(* IEC 61131-3 sources: ControlsBenchMUSE/codesys/demo/source, 10 files *)

(* ---- ST_BenchInputImage.st ---- *)
TYPE ST_BenchInputImage :
STRUCT
    PE_Entry : BOOL;
    PE_D1Approach : BOOL;
    PE_D2Approach : BOOL;
    PE_ExitA : BOOL;
    PE_ExitB : BOOL;
    PE_Runout : BOOL;
    D1_HomeFB : BOOL;
    D1_ExtendedFB : BOOL;
    D2_HomeFB : BOOL;
    D2_ExtendedFB : BOOL;
    Drive_RunningFB : BOOL;
    Drive_Overload : BOOL;
    ExitA_Ready : BOOL;
    ExitB_Ready : BOOL;
    Runout_Ready : BOOL;
    Belt_SpeedActual : REAL;
    Drive_Current : REAL;
    D1_Position : REAL;
    D2_Position : REAL;
    Encoder_Count : UDINT;
END_STRUCT
END_TYPE

(* ---- ST_DemoStatus.st ---- *)
TYPE ST_DemoStatus :
STRUCT
    Mode : UINT;
    ModeText : STRING(16);
    FaultCode : UINT;
    FaultText : STRING(80);
    ExceptionCode : UINT;
    ExceptionText : STRING(80);
    Motor_RunCmd : BOOL;
    D1_ExtendCmd : BOOL;
    D2_ExtendCmd : BOOL;
    StackLight_Red : BOOL;
    StackLight_Green : BOOL;
    ReleaseReady : BOOL;
    ItemActive : BOOL;
    ActiveItemId : UDINT;
    RequestedRoute : UINT;
    EffectiveRoute : UINT;
    ActualExit : UINT;
    Disposition : UINT;
    OfferAckSequence : UDINT;
    OfferAckItemId : UDINT;
    OfferAccepted : BOOL;
    OfferReason : UINT;
    OfferPending : BOOL;
    CompletionSequence : UDINT;
    CompletionPending : BOOL;
    CompletionItemId : UDINT;
    CompletionRoute : UINT;
    CompletionExit : UINT;
    CompletionDisposition : UINT;
    CountExitA : UDINT;
    CountExitB : UDINT;
    CountRunout : UDINT;
    CountMisroute : UDINT;
    CountFaulted : UDINT;
    StartAck : UDINT;
    StopAck : UDINT;
    ResetAck : UDINT;
    StartAccepted : BOOL;
    ResetAccepted : BOOL;
    EncoderDelta : UDINT;
    BeltSpeedMps : LREAL;
    TravelMetres : LREAL;
    ScanTimeUs : ULINT;
END_STRUCT
END_TYPE

(* ---- GVL_BenchRead.st ---- *)
NAMESPACE GVL_BenchRead
{attribute 'qualified_only'}
VAR_GLOBAL
    // Bench state and liveness. Workstation read-only through OPC UA.
    SimApplied : BOOL := FALSE;
    ConnectorStale : BOOL := TRUE;
    ActiveSlot : USINT := 255;
    AppliedEpoch : ULINT := 0;
    AppliedSequence : ULINT := 0;
    // Published compatibility placeholders retained by the configured symbol type.
    AppliedCaptureCycle : ULINT := 0;
    AppliedCaptureTimeUs : ULINT := 0;
    PlcHeartbeat : ULINT := 0;
    PlcBootIdentity : ULINT := 0;
    PlcCycle : ULINT := 0;
    PlcTimeUs : ULINT := 0;

    // Commit diagnostics.
    AppliedCommitCount : ULINT := 0;
    DuplicateCommitCount : ULINT := 0;
    StaleCommitCount : ULINT := 0;
    SkippedSequenceCount : ULINT := 0;
    InvalidSlotCount : ULINT := 0;
    InvalidPayloadCount : ULINT := 0;
    SlotMetadataMismatchCount : ULINT := 0;
    EpochRejectedCount : ULINT := 0;
    SessionResetCount : ULINT := 0;

    // Application-visible active raw input image.
    Active_PE_Entry : BOOL := FALSE;
    Active_PE_D1Approach : BOOL := FALSE;
    Active_PE_D2Approach : BOOL := FALSE;
    Active_PE_ExitA : BOOL := FALSE;
    Active_PE_ExitB : BOOL := FALSE;
    Active_PE_Runout : BOOL := FALSE;
    Active_D1_HomeFB : BOOL := FALSE;
    Active_D1_ExtendedFB : BOOL := FALSE;
    Active_D2_HomeFB : BOOL := FALSE;
    Active_D2_ExtendedFB : BOOL := FALSE;
    Active_Drive_RunningFB : BOOL := FALSE;
    Active_Drive_Overload : BOOL := FALSE;
    Active_ExitA_Ready : BOOL := FALSE;
    Active_ExitB_Ready : BOOL := FALSE;
    Active_Runout_Ready : BOOL := FALSE;
    Active_Belt_SpeedActual : REAL := 0.0;
    Active_Drive_Current : REAL := 0.0;
    Active_D1_Position : REAL := 0.0;
    Active_D2_Position : REAL := 0.0;
    Active_Encoder_Count : UDINT := 0;

    // Fixture-only deterministic PLC output image.
    Motor_RunCmd : BOOL := FALSE;
    D1_ExtendCmd : BOOL := FALSE;
    D2_ExtendCmd : BOOL := FALSE;
    StackLight_Red : BOOL := FALSE;
    StackLight_Green : BOOL := FALSE;
    OutputSourceEpoch : ULINT := 0;
    OutputSourceSequence : ULINT := 0;
    OutputSourceAppliedCycle : ULINT := 0;
    OutputCaptureCycle : ULINT := 0;
    OutputCaptureTimeUs : ULINT := 0;
END_VAR
END_NAMESPACE

(* ---- GVL_BenchWrite.st ---- *)
NAMESPACE GVL_BenchWrite
{attribute 'qualified_only'}
VAR_GLOBAL
    // Bench authority and commit request. Workstation-writable through OPC UA.
    SimRequest : BOOL := FALSE;
    SessionResetRequest : BOOL := FALSE;
    RequestedSlot : USINT := 0;
    RequestedEpoch : ULINT := 0;
    RequestedSequence : ULINT := 0;
    // Published compatibility placeholder; RequestedSequence is the active commit edge.
    CommitToken : ULINT := 0;
    WorkstationHeartbeat : ULINT := 0;

    // Slot 0 metadata.
    Slot0_Valid : BOOL := FALSE;
    Slot0_Epoch : ULINT := 0;
    Slot0_Sequence : ULINT := 0;

    // Slot 0 complete raw input image.
    Slot0_PE_Entry : BOOL := FALSE;
    Slot0_PE_D1Approach : BOOL := FALSE;
    Slot0_PE_D2Approach : BOOL := FALSE;
    Slot0_PE_ExitA : BOOL := FALSE;
    Slot0_PE_ExitB : BOOL := FALSE;
    Slot0_PE_Runout : BOOL := FALSE;
    Slot0_D1_HomeFB : BOOL := FALSE;
    Slot0_D1_ExtendedFB : BOOL := FALSE;
    Slot0_D2_HomeFB : BOOL := FALSE;
    Slot0_D2_ExtendedFB : BOOL := FALSE;
    Slot0_Drive_RunningFB : BOOL := FALSE;
    Slot0_Drive_Overload : BOOL := FALSE;
    Slot0_ExitA_Ready : BOOL := FALSE;
    Slot0_ExitB_Ready : BOOL := FALSE;
    Slot0_Runout_Ready : BOOL := FALSE;
    Slot0_Belt_SpeedActual : REAL := 0.0;
    Slot0_Drive_Current : REAL := 0.0;
    Slot0_D1_Position : REAL := 0.0;
    Slot0_D2_Position : REAL := 0.0;
    Slot0_Encoder_Count : UDINT := 0;

    // Slot 1 metadata.
    Slot1_Valid : BOOL := FALSE;
    Slot1_Epoch : ULINT := 0;
    Slot1_Sequence : ULINT := 0;

    // Slot 1 complete raw input image.
    Slot1_PE_Entry : BOOL := FALSE;
    Slot1_PE_D1Approach : BOOL := FALSE;
    Slot1_PE_D2Approach : BOOL := FALSE;
    Slot1_PE_ExitA : BOOL := FALSE;
    Slot1_PE_ExitB : BOOL := FALSE;
    Slot1_PE_Runout : BOOL := FALSE;
    Slot1_D1_HomeFB : BOOL := FALSE;
    Slot1_D1_ExtendedFB : BOOL := FALSE;
    Slot1_D2_HomeFB : BOOL := FALSE;
    Slot1_D2_ExtendedFB : BOOL := FALSE;
    Slot1_Drive_RunningFB : BOOL := FALSE;
    Slot1_Drive_Overload : BOOL := FALSE;
    Slot1_ExitA_Ready : BOOL := FALSE;
    Slot1_ExitB_Ready : BOOL := FALSE;
    Slot1_Runout_Ready : BOOL := FALSE;
    Slot1_Belt_SpeedActual : REAL := 0.0;
    Slot1_Drive_Current : REAL := 0.0;
    Slot1_D1_Position : REAL := 0.0;
    Slot1_D2_Position : REAL := 0.0;
    Slot1_Encoder_Count : UDINT := 0;
END_VAR
END_NAMESPACE

(* ---- GVL_DemoHardware.st ---- *)
NAMESPACE GVL_DemoHardware
{attribute 'qualified_only'}
VAR_GLOBAL
    // Physical adapter boundary; map hardware acquisition here. No hardware on Control Win.
    Inputs : ST_BenchInputImage;
    Motor_RunCmd : BOOL;
    D1_ExtendCmd : BOOL;
    D2_ExtendCmd : BOOL;
    StackLight_Red : BOOL;
    StackLight_Green : BOOL;
END_VAR
END_NAMESPACE

(* ---- GVL_DemoRead.st ---- *)
NAMESPACE GVL_DemoRead
{attribute 'qualified_only'}
VAR_GLOBAL
    BuildId : UDINT := 8001;
    InterfaceVersion : UINT := 1;
    Status : ST_DemoStatus;
END_VAR
END_NAMESPACE

(* ---- GVL_DemoWrite.st ---- *)
NAMESPACE GVL_DemoWrite
{attribute 'qualified_only'}
VAR_GLOBAL
    StartSequence : UDINT := 0;
    StopSequence : UDINT := 0;
    ResetSequence : UDINT := 0;
    AutoRequest : BOOL := FALSE;
    OfferSequence : UDINT := 0;
    OfferItemId : UDINT := 0;
    OfferRoute : UINT := 0;
    CompletionAck : UDINT := 0;
END_VAR
END_NAMESPACE

(* ---- FB_BenchIntercept.st ---- *)
FUNCTION_BLOCK FB_BenchIntercept
VAR_INPUT
    Hardware : ST_BenchInputImage;
END_VAR
VAR_OUTPUT
    Image : ST_BenchInputImage;
END_VAR
VAR
    previousSim : BOOL;
    simulationEntry : BOOL;
    ActiveImage : ST_BenchInputImage;
    CandidateImage : ST_BenchInputImage;
    ZeroImage : ST_BenchInputImage;

    initialized : BOOL := FALSE;
    haveHeartbeat : BOOL := FALSE;
    previousSessionReset : BOOL := FALSE;
    lastWorkstationHeartbeat : ULINT := 0;
    lastHeartbeatCycle : ULINT := 0;

    lastRequestSequence : ULINT := 0;

    requestChanged : BOOL;
    sessionResetEdge : BOOL;
    slotIsInactive : BOOL;
    slotValid : BOOL;
    slotEpoch : ULINT;
    slotSequence : ULINT;
    acceptCommit : BOOL;
    payloadPhysicalValid : BOOL;

    nowUs : SysTimeCore.SYSTIME;
    timeResult : UDINT;
END_VAR
// Capture monotonic PLC time and advance scan-owned liveness.
timeResult := SysTimeCore.SysTimeGetUs(nowUs);
GVL_BenchRead.PlcTimeUs := nowUs;
GVL_BenchRead.PlcCycle := GVL_BenchRead.PlcCycle + 1;
GVL_BenchRead.PlcHeartbeat := GVL_BenchRead.PlcHeartbeat + 1;

IF NOT initialized THEN
    GVL_BenchRead.PlcBootIdentity := nowUs;
    IF GVL_BenchRead.PlcBootIdentity = 0 THEN
        GVL_BenchRead.PlcBootIdentity := 1;
    END_IF;
    GVL_BenchRead.ActiveSlot := 255;
    ActiveImage := ZeroImage;
    initialized := TRUE;
END_IF;

// Hardware passthrough is the cold-start default. Entering simulation zeros all raw types.
simulationEntry := GVL_BenchWrite.SimRequest AND NOT previousSim;
previousSim := GVL_BenchWrite.SimRequest;
GVL_BenchRead.SimApplied := GVL_BenchWrite.SimRequest;
IF simulationEntry THEN
    ActiveImage := ZeroImage;
    GVL_BenchRead.AppliedEpoch := 0;
    GVL_BenchRead.AppliedSequence := 0;
    GVL_BenchRead.ActiveSlot := 255;
    lastRequestSequence := GVL_BenchWrite.RequestedSequence;
END_IF;

// Heartbeat freshness is independent of commit traffic.
// 25 scans at the current 20 ms task interval equals the 500 ms M5 floor.
IF GVL_BenchWrite.WorkstationHeartbeat <> lastWorkstationHeartbeat THEN
    lastWorkstationHeartbeat := GVL_BenchWrite.WorkstationHeartbeat;
    lastHeartbeatCycle := GVL_BenchRead.PlcCycle;
    haveHeartbeat := TRUE;
END_IF;

IF haveHeartbeat THEN
    GVL_BenchRead.ConnectorStale :=
        (GVL_BenchRead.PlcCycle - lastHeartbeatCycle) > 25;
ELSE
    GVL_BenchRead.ConnectorStale := TRUE;
END_IF;

// A rising session reset explicitly clears epoch continuity and the active image.
sessionResetEdge :=
    GVL_BenchWrite.SessionResetRequest AND NOT previousSessionReset;
previousSessionReset := GVL_BenchWrite.SessionResetRequest;

IF sessionResetEdge THEN
    GVL_BenchRead.AppliedEpoch := 0;
    GVL_BenchRead.AppliedSequence := 0;
    GVL_BenchRead.ActiveSlot := 255;
    ActiveImage := ZeroImage;
    lastRequestSequence := GVL_BenchWrite.RequestedSequence;
    GVL_BenchRead.SessionResetCount :=
        GVL_BenchRead.SessionResetCount + 1;
END_IF;

// RequestedSequence is the single commit edge and is written after the complete valid slot.
requestChanged := GVL_BenchWrite.RequestedSequence <> lastRequestSequence;

IF GVL_BenchRead.SimApplied
    AND NOT sessionResetEdge
    AND requestChanged
    AND ((GVL_BenchWrite.RequestedEpoch <> 0)
        OR (GVL_BenchWrite.RequestedSequence <> 0)) THEN

    acceptCommit := FALSE;
    slotValid := FALSE;
    slotEpoch := 0;
    slotSequence := 0;

    IF GVL_BenchWrite.RequestedSlot > 1 THEN
        GVL_BenchRead.InvalidSlotCount :=
            GVL_BenchRead.InvalidSlotCount + 1;
    ELSE
        slotIsInactive :=
            (GVL_BenchRead.ActiveSlot = 255)
            OR (GVL_BenchWrite.RequestedSlot <> GVL_BenchRead.ActiveSlot);

        IF NOT slotIsInactive THEN
            GVL_BenchRead.InvalidSlotCount :=
                GVL_BenchRead.InvalidSlotCount + 1;
        ELSE
            IF GVL_BenchWrite.RequestedSlot = 0 THEN
                slotValid := GVL_BenchWrite.Slot0_Valid;
                slotEpoch := GVL_BenchWrite.Slot0_Epoch;
                slotSequence := GVL_BenchWrite.Slot0_Sequence;

                CandidateImage.PE_Entry := GVL_BenchWrite.Slot0_PE_Entry;
                CandidateImage.PE_D1Approach := GVL_BenchWrite.Slot0_PE_D1Approach;
                CandidateImage.PE_D2Approach := GVL_BenchWrite.Slot0_PE_D2Approach;
                CandidateImage.PE_ExitA := GVL_BenchWrite.Slot0_PE_ExitA;
                CandidateImage.PE_ExitB := GVL_BenchWrite.Slot0_PE_ExitB;
                CandidateImage.PE_Runout := GVL_BenchWrite.Slot0_PE_Runout;
                CandidateImage.D1_HomeFB := GVL_BenchWrite.Slot0_D1_HomeFB;
                CandidateImage.D1_ExtendedFB := GVL_BenchWrite.Slot0_D1_ExtendedFB;
                CandidateImage.D2_HomeFB := GVL_BenchWrite.Slot0_D2_HomeFB;
                CandidateImage.D2_ExtendedFB := GVL_BenchWrite.Slot0_D2_ExtendedFB;
                CandidateImage.Drive_RunningFB := GVL_BenchWrite.Slot0_Drive_RunningFB;
                CandidateImage.Drive_Overload := GVL_BenchWrite.Slot0_Drive_Overload;
                CandidateImage.ExitA_Ready := GVL_BenchWrite.Slot0_ExitA_Ready;
                CandidateImage.ExitB_Ready := GVL_BenchWrite.Slot0_ExitB_Ready;
                CandidateImage.Runout_Ready := GVL_BenchWrite.Slot0_Runout_Ready;
                CandidateImage.Belt_SpeedActual := GVL_BenchWrite.Slot0_Belt_SpeedActual;
                CandidateImage.Drive_Current := GVL_BenchWrite.Slot0_Drive_Current;
                CandidateImage.D1_Position := GVL_BenchWrite.Slot0_D1_Position;
                CandidateImage.D2_Position := GVL_BenchWrite.Slot0_D2_Position;
                CandidateImage.Encoder_Count := GVL_BenchWrite.Slot0_Encoder_Count;
            ELSE
                slotValid := GVL_BenchWrite.Slot1_Valid;
                slotEpoch := GVL_BenchWrite.Slot1_Epoch;
                slotSequence := GVL_BenchWrite.Slot1_Sequence;

                CandidateImage.PE_Entry := GVL_BenchWrite.Slot1_PE_Entry;
                CandidateImage.PE_D1Approach := GVL_BenchWrite.Slot1_PE_D1Approach;
                CandidateImage.PE_D2Approach := GVL_BenchWrite.Slot1_PE_D2Approach;
                CandidateImage.PE_ExitA := GVL_BenchWrite.Slot1_PE_ExitA;
                CandidateImage.PE_ExitB := GVL_BenchWrite.Slot1_PE_ExitB;
                CandidateImage.PE_Runout := GVL_BenchWrite.Slot1_PE_Runout;
                CandidateImage.D1_HomeFB := GVL_BenchWrite.Slot1_D1_HomeFB;
                CandidateImage.D1_ExtendedFB := GVL_BenchWrite.Slot1_D1_ExtendedFB;
                CandidateImage.D2_HomeFB := GVL_BenchWrite.Slot1_D2_HomeFB;
                CandidateImage.D2_ExtendedFB := GVL_BenchWrite.Slot1_D2_ExtendedFB;
                CandidateImage.Drive_RunningFB := GVL_BenchWrite.Slot1_Drive_RunningFB;
                CandidateImage.Drive_Overload := GVL_BenchWrite.Slot1_Drive_Overload;
                CandidateImage.ExitA_Ready := GVL_BenchWrite.Slot1_ExitA_Ready;
                CandidateImage.ExitB_Ready := GVL_BenchWrite.Slot1_ExitB_Ready;
                CandidateImage.Runout_Ready := GVL_BenchWrite.Slot1_Runout_Ready;
                CandidateImage.Belt_SpeedActual := GVL_BenchWrite.Slot1_Belt_SpeedActual;
                CandidateImage.Drive_Current := GVL_BenchWrite.Slot1_Drive_Current;
                CandidateImage.D1_Position := GVL_BenchWrite.Slot1_D1_Position;
                CandidateImage.D2_Position := GVL_BenchWrite.Slot1_D2_Position;
                CandidateImage.Encoder_Count := GVL_BenchWrite.Slot1_Encoder_Count;
            END_IF;

            // Generous fixture limits reject NaN, infinity, and physically invalid negatives.
            payloadPhysicalValid :=
                (CandidateImage.Belt_SpeedActual >= 0.0)
                AND (CandidateImage.Belt_SpeedActual <= 100.0)
                AND (CandidateImage.Drive_Current >= 0.0)
                AND (CandidateImage.Drive_Current <= 10000.0)
                AND (CandidateImage.D1_Position >= 0.0)
                AND (CandidateImage.D1_Position <= 100.0)
                AND (CandidateImage.D2_Position >= 0.0)
                AND (CandidateImage.D2_Position <= 100.0);

            IF NOT slotValid THEN
                GVL_BenchRead.InvalidPayloadCount :=
                    GVL_BenchRead.InvalidPayloadCount + 1;
            ELSIF NOT payloadPhysicalValid THEN
                GVL_BenchRead.InvalidPayloadCount :=
                    GVL_BenchRead.InvalidPayloadCount + 1;
            ELSIF (slotEpoch = 0) OR (slotSequence = 0) THEN
                GVL_BenchRead.InvalidPayloadCount :=
                    GVL_BenchRead.InvalidPayloadCount + 1;
            ELSIF (slotEpoch <> GVL_BenchWrite.RequestedEpoch)
                OR (slotSequence <> GVL_BenchWrite.RequestedSequence) THEN
                GVL_BenchRead.SlotMetadataMismatchCount :=
                    GVL_BenchRead.SlotMetadataMismatchCount + 1;
            ELSIF GVL_BenchRead.AppliedEpoch = 0 THEN
                acceptCommit := TRUE;
            ELSIF slotEpoch = GVL_BenchRead.AppliedEpoch THEN
                IF slotSequence = GVL_BenchRead.AppliedSequence THEN
                    GVL_BenchRead.DuplicateCommitCount :=
                        GVL_BenchRead.DuplicateCommitCount + 1;
                ELSIF slotSequence < GVL_BenchRead.AppliedSequence THEN
                    GVL_BenchRead.StaleCommitCount :=
                        GVL_BenchRead.StaleCommitCount + 1;
                ELSE
                    IF slotSequence > (GVL_BenchRead.AppliedSequence + 1) THEN
                        GVL_BenchRead.SkippedSequenceCount :=
                            GVL_BenchRead.SkippedSequenceCount + 1;
                    END_IF;
                    acceptCommit := TRUE;
                END_IF;
            ELSIF GVL_BenchRead.ConnectorStale OR sessionResetEdge THEN
                // A new random workstation epoch is allowed only after stale or explicit reset.
                acceptCommit := TRUE;
            ELSE
                GVL_BenchRead.EpochRejectedCount :=
                    GVL_BenchRead.EpochRejectedCount + 1;
            END_IF;

            IF acceptCommit THEN
                // Same-task scan-owned publication: downstream logic sees one complete revision.
                ActiveImage := CandidateImage;
                GVL_BenchRead.ActiveSlot := GVL_BenchWrite.RequestedSlot;
                GVL_BenchRead.AppliedEpoch := slotEpoch;
                GVL_BenchRead.AppliedSequence := slotSequence;
                GVL_BenchRead.AppliedCaptureCycle := GVL_BenchRead.PlcCycle;
                GVL_BenchRead.AppliedCaptureTimeUs := GVL_BenchRead.PlcTimeUs;
                GVL_BenchRead.AppliedCommitCount :=
                    GVL_BenchRead.AppliedCommitCount + 1;
            END_IF;
        END_IF;
    END_IF;

END_IF;

IF requestChanged THEN
    lastRequestSequence := GVL_BenchWrite.RequestedSequence;
END_IF;

// Select the complete image before any application logic executes.
IF GVL_BenchRead.SimApplied THEN
    Image := ActiveImage;
ELSE
    Image := Hardware;
END_IF;
// Publish the selected application-visible raw image for verification.
GVL_BenchRead.Active_PE_Entry := Image.PE_Entry;
GVL_BenchRead.Active_PE_D1Approach := Image.PE_D1Approach;
GVL_BenchRead.Active_PE_D2Approach := Image.PE_D2Approach;
GVL_BenchRead.Active_PE_ExitA := Image.PE_ExitA;
GVL_BenchRead.Active_PE_ExitB := Image.PE_ExitB;
GVL_BenchRead.Active_PE_Runout := Image.PE_Runout;
GVL_BenchRead.Active_D1_HomeFB := Image.D1_HomeFB;
GVL_BenchRead.Active_D1_ExtendedFB := Image.D1_ExtendedFB;
GVL_BenchRead.Active_D2_HomeFB := Image.D2_HomeFB;
GVL_BenchRead.Active_D2_ExtendedFB := Image.D2_ExtendedFB;
GVL_BenchRead.Active_Drive_RunningFB := Image.Drive_RunningFB;
GVL_BenchRead.Active_Drive_Overload := Image.Drive_Overload;
GVL_BenchRead.Active_ExitA_Ready := Image.ExitA_Ready;
GVL_BenchRead.Active_ExitB_Ready := Image.ExitB_Ready;
GVL_BenchRead.Active_Runout_Ready := Image.Runout_Ready;
GVL_BenchRead.Active_Belt_SpeedActual := Image.Belt_SpeedActual;
GVL_BenchRead.Active_Drive_Current := Image.Drive_Current;
GVL_BenchRead.Active_D1_Position := Image.D1_Position;
GVL_BenchRead.Active_D2_Position := Image.D2_Position;
GVL_BenchRead.Active_Encoder_Count := Image.Encoder_Count;
END_FUNCTION_BLOCK

(* ---- FB_DemoConveyor.st ---- *)
FUNCTION_BLOCK FB_DemoConveyor
VAR_INPUT
    I : ST_BenchInputImage;
    NowUs : ULINT;
    StartSequence : UDINT;
    StopSequence : UDINT;
    ResetSequence : UDINT;
    AutoRequest : BOOL;
    OfferSequence : UDINT;
    OfferItemId : UDINT;
    OfferRoute : UINT;
    CompletionAck : UDINT;
END_VAR
VAR_OUTPUT
    Q : ST_DemoStatus;
END_VAR
VAR
    prev : ST_BenchInputImage;
    initialized : BOOL;
    encoderPrevious : UDINT;
    speedCounts : ULINT;
    speedStartUs : ULINT;
    previousStart : UDINT;
    previousStop : UDINT;
    previousReset : UDINT;
    previousOffer : UDINT;
    pendingId : UDINT;
    pendingRoute : UINT;
    passedD1 : BOOL;
    passedD2 : BOOL;
    runningSeen : BOOL;
    startEdge : BOOL;
    stopEdge : BOOL;
    resetEdge : BOOL;
    entryEdge : BOOL;
    exitAEdge : BOOL;
    exitBEdge : BOOL;
    runoutEdge : BOOL;
    exitEdges : UINT;
    clearBeams : BOOL;
    readyToStart : BOOL;
    readyToResume : BOOL;
    observedExit : UINT;
    observedDisposition : UINT;
    tMotorStart : TON;
    tMotorLost : TON;
    tStop : TON;
    tStill : TON;
    tD1Extend : TON;
    tD2Extend : TON;
    tD1Home : TON;
    tD2Home : TON;
    tTransit : TON;
END_VAR
// Raw counter scaling stays inside the actual PLC, including UDINT rollover.
IF NOT initialized THEN
    encoderPrevious := I.Encoder_Count;
    speedStartUs := NowUs;
    initialized := TRUE;
END_IF;
IF I.Encoder_Count >= encoderPrevious THEN
    Q.EncoderDelta := I.Encoder_Count - encoderPrevious;
ELSE
    Q.EncoderDelta := ULINT_TO_UDINT(ULINT#4294967296 - UDINT_TO_ULINT(encoderPrevious)
        + UDINT_TO_ULINT(I.Encoder_Count));
END_IF;
encoderPrevious := I.Encoder_Count;
speedCounts := speedCounts + UDINT_TO_ULINT(Q.EncoderDelta);
Q.TravelMetres := Q.TravelMetres + UDINT_TO_LREAL(Q.EncoderDelta) / 1000.0;
IF NowUs - speedStartUs >= 100000 THEN
    Q.BeltSpeedMps := ULINT_TO_LREAL(speedCounts) * 1000.0 / ULINT_TO_LREAL(NowUs - speedStartUs);
    speedCounts := 0;
    speedStartUs := NowUs;
END_IF;
Q.ScanTimeUs := NowUs;

startEdge := StartSequence <> previousStart;
stopEdge := StopSequence <> previousStop;
resetEdge := ResetSequence <> previousReset;
previousStart := StartSequence;
previousStop := StopSequence;
previousReset := ResetSequence;
entryEdge := I.PE_Entry AND NOT prev.PE_Entry;
exitAEdge := I.PE_ExitA AND NOT prev.PE_ExitA;
exitBEdge := I.PE_ExitB AND NOT prev.PE_ExitB;
runoutEdge := I.PE_Runout AND NOT prev.PE_Runout;
exitEdges := BOOL_TO_UINT(exitAEdge) + BOOL_TO_UINT(exitBEdge) + BOOL_TO_UINT(runoutEdge);
clearBeams := NOT (I.PE_Entry OR I.PE_D1Approach OR I.PE_D2Approach
    OR I.PE_ExitA OR I.PE_ExitB OR I.PE_Runout);
Q.CompletionPending := Q.CompletionSequence <> CompletionAck;

// Offers use an immutable payload followed by a write-last sequence. Duplicate sequences do nothing.
IF (OfferSequence <> 0) AND (OfferSequence < previousOffer) THEN
    Q.OfferAckSequence := OfferSequence;
    Q.OfferAckItemId := OfferItemId;
    Q.OfferAccepted := FALSE;
    Q.OfferReason := 4; // stale/replayed sequence; never enqueue again
END_IF;
IF OfferSequence > previousOffer THEN
    previousOffer := OfferSequence;
    Q.OfferAckSequence := OfferSequence;
    Q.OfferAckItemId := OfferItemId;
    Q.OfferAccepted := FALSE;
    Q.OfferReason := 1; // busy/unavailable
    IF (OfferRoute > 2) OR (OfferItemId = 0) THEN
        Q.OfferReason := 2; // malformed
    ELSIF (Q.Mode <> 3) AND NOT Q.CompletionPending THEN
        IF Q.ItemActive THEN
            IF ((Q.ActiveItemId = 0) OR (Q.ActiveItemId = OfferItemId))
                AND ((Q.RequestedRoute = 0) OR (Q.RequestedRoute = OfferRoute)) THEN
                Q.ActiveItemId := OfferItemId;
                Q.RequestedRoute := OfferRoute;
                Q.OfferAccepted := TRUE;
                Q.OfferReason := 0;
            ELSE
                Q.OfferReason := 3; // conflicting identity/assignment
            END_IF;
        ELSIF NOT Q.OfferPending THEN
            pendingId := OfferItemId;
            pendingRoute := OfferRoute;
            Q.OfferPending := TRUE;
            Q.OfferAccepted := TRUE;
            Q.OfferReason := 0;
        END_IF;
    END_IF;
END_IF;

// Stop and Auto withdrawal both remove the run command in this scan.
IF stopEdge THEN Q.StopAck := StopSequence; END_IF;
IF (stopEdge OR NOT AutoRequest) AND (Q.Mode = 1) THEN Q.Mode := 2; END_IF;

readyToStart := NOT I.Drive_Overload
    AND I.D1_HomeFB AND NOT I.D1_ExtendedFB
    AND I.D2_HomeFB AND NOT I.D2_ExtendedFB
    AND I.Runout_Ready;
readyToResume := Q.ItemActive AND NOT I.Drive_Overload AND I.Runout_Ready
    AND ((I.D1_HomeFB AND NOT I.D1_ExtendedFB)
        OR ((Q.EffectiveRoute = 1) AND I.D1_ExtendedFB AND NOT I.D1_HomeFB))
    AND ((I.D2_HomeFB AND NOT I.D2_ExtendedFB)
        OR ((Q.EffectiveRoute = 2) AND I.D2_ExtendedFB AND NOT I.D2_HomeFB));
IF resetEdge THEN
    Q.ResetAck := ResetSequence;
    Q.ResetAccepted := FALSE;
    IF (Q.Mode <> 1) AND (Q.Mode <> 2) AND readyToStart
        AND NOT I.Drive_RunningFB AND clearBeams AND NOT Q.CompletionPending THEN
        Q.FaultCode := 0;
        Q.FaultText := '';
        Q.ExceptionCode := 0;
        Q.ExceptionText := '';
        Q.OfferPending := FALSE;
        Q.Mode := 0;
        runningSeen := FALSE;
        Q.ResetAccepted := TRUE;
    END_IF;
END_IF;
IF startEdge THEN
    Q.StartAck := StartSequence;
    Q.StartAccepted := FALSE;
    IF (Q.Mode = 0) AND AutoRequest AND (readyToStart OR readyToResume) AND NOT stopEdge
        AND NOT Q.CompletionPending AND (clearBeams OR Q.ItemActive) THEN
        Q.Mode := 1;
        runningSeen := FALSE;
        Q.StartAccepted := TRUE;
    END_IF;
END_IF;

// Accept one physical carton. A second carton is outside this baseline capacity.
IF entryEdge THEN
    IF Q.ItemActive OR Q.CompletionPending OR (Q.Mode <> 1) OR NOT I.Drive_RunningFB THEN
        Trip(Code := 30, Text := 'Unexpected entry / single-carton capacity exceeded');
    ELSE
        Q.ItemActive := TRUE;
        Q.ActiveItemId := 0;
        Q.RequestedRoute := 0;
        IF Q.OfferPending THEN
            Q.ActiveItemId := pendingId;
            Q.RequestedRoute := pendingRoute;
            Q.OfferPending := FALSE;
        END_IF;
        Q.EffectiveRoute := 0;
        Q.ActualExit := 0;
        Q.Disposition := 0;
        Q.ExceptionCode := 0;
        Q.ExceptionText := '';
        passedD1 := FALSE;
        passedD2 := FALSE;
    END_IF;
END_IF;

// Preposition as soon as an assignment exists. Each approach edge locks reachability.
IF Q.ItemActive THEN
    IF NOT passedD1 AND NOT passedD2 THEN
        Q.EffectiveRoute := 0;
        IF (Q.RequestedRoute = 1) AND I.ExitA_Ready THEN Q.EffectiveRoute := 1; END_IF;
        IF (Q.RequestedRoute = 2) AND I.ExitB_Ready THEN Q.EffectiveRoute := 2; END_IF;
    ELSIF NOT passedD2 AND (Q.EffectiveRoute <> 1) THEN
        Q.EffectiveRoute := 0;
        IF (Q.RequestedRoute = 2) AND I.ExitB_Ready THEN Q.EffectiveRoute := 2; END_IF;
    END_IF;
    IF I.PE_D1Approach AND NOT prev.PE_D1Approach THEN passedD1 := TRUE; END_IF;
    IF I.PE_D2Approach AND NOT prev.PE_D2Approach THEN passedD2 := TRUE; END_IF;
    IF (Q.RequestedRoute <> 0) AND (Q.EffectiveRoute = 0) THEN
        Q.ExceptionCode := 1;
        Q.ExceptionText := 'Assigned route unavailable or received too late; runout';
    END_IF;
END_IF;
Q.Motor_RunCmd := Q.Mode = 1;
Q.D1_ExtendCmd := Q.ItemActive AND (Q.EffectiveRoute = 1) AND (Q.Mode <> 3);
Q.D2_ExtendCmd := Q.ItemActive AND (Q.EffectiveRoute = 2) AND (Q.Mode <> 3);

IF (Q.Mode = 1) AND I.Drive_RunningFB THEN runningSeen := TRUE; END_IF;
tMotorStart(IN := (Q.Mode = 1) AND NOT runningSeen AND NOT I.Drive_RunningFB, PT := T#1500ms);
tMotorLost(IN := (Q.Mode = 1) AND runningSeen AND NOT I.Drive_RunningFB, PT := T#500ms);
tStill(IN := NOT I.Drive_RunningFB AND (Q.EncoderDelta = 0), PT := T#200ms);
tStop(IN := (Q.Mode = 2) AND NOT tStill.Q, PT := T#4s);
tD1Extend(IN := Q.D1_ExtendCmd AND NOT I.D1_ExtendedFB, PT := T#1200ms);
tD2Extend(IN := Q.D2_ExtendCmd AND NOT I.D2_ExtendedFB, PT := T#1200ms);
tD1Home(IN := (Q.Mode = 1 OR Q.Mode = 2) AND NOT Q.D1_ExtendCmd AND NOT I.D1_HomeFB, PT := T#1200ms);
tD2Home(IN := (Q.Mode = 1 OR Q.Mode = 2) AND NOT Q.D2_ExtendCmd AND NOT I.D2_HomeFB, PT := T#1200ms);
tTransit(IN := Q.ItemActive AND (Q.Mode = 1), PT := T#30s);

// Machine faults take priority over exit success in the same scan.
IF I.Drive_Overload THEN Trip(Code := 10, Text := 'Drive overload'); END_IF;
IF I.D1_HomeFB AND I.D1_ExtendedFB THEN Trip(Code := 21, Text := 'D1 contradictory limits'); END_IF;
IF I.D2_HomeFB AND I.D2_ExtendedFB THEN Trip(Code := 22, Text := 'D2 contradictory limits'); END_IF;
IF tMotorStart.Q THEN Trip(Code := 11, Text := 'Motor running feedback missing on start'); END_IF;
IF tMotorLost.Q THEN Trip(Code := 12, Text := 'Motor running feedback lost'); END_IF;
IF tStop.Q THEN Trip(Code := 13, Text := 'Motor failed to stop within 4 seconds'); END_IF;
IF tD1Extend.Q THEN Trip(Code := 23, Text := 'D1 extend feedback timeout'); END_IF;
IF tD2Extend.Q THEN Trip(Code := 24, Text := 'D2 extend feedback timeout'); END_IF;
IF tD1Home.Q THEN Trip(Code := 25, Text := 'D1 home feedback timeout'); END_IF;
IF tD2Home.Q THEN Trip(Code := 26, Text := 'D2 home feedback timeout'); END_IF;
IF tTransit.Q THEN Trip(Code := 33, Text := 'Carton transit timeout'); END_IF;
IF (Q.Mode = 1) AND NOT I.Runout_Ready THEN Trip(Code := 34, Text := 'Runout unavailable; conveyor stopped'); END_IF;
IF exitEdges > 1 THEN Trip(Code := 31, Text := 'Multiple exit edges for single carton'); END_IF;
IF (exitEdges = 1) AND (Q.Mode <> 3) THEN
    IF Q.ItemActive THEN
        observedExit := 3;
        IF exitAEdge THEN observedExit := 1; END_IF;
        IF exitBEdge THEN observedExit := 2; END_IF;
        observedDisposition := 3; // misroute
        IF Q.RequestedRoute = observedExit THEN observedDisposition := 1; END_IF;
        IF (Q.RequestedRoute = 0) AND (observedExit = 3) THEN observedDisposition := 2; END_IF;
        IF (observedDisposition = 1) AND
            (((observedExit = 1) AND (NOT I.D1_ExtendedFB OR I.D1_HomeFB))
            OR ((observedExit = 2) AND (NOT I.D2_ExtendedFB OR I.D2_HomeFB))) THEN
            Trip(Code := 27, Text := 'Assigned exit observed without verified divert position');
        ELSE
            Finish(Actual := observedExit, Result := observedDisposition);
        END_IF;
    ELSE
        Trip(Code := 32, Text := 'Exit without an active tracked carton');
    END_IF;
END_IF;

IF (Q.Mode = 2) AND tStill.Q THEN Q.Mode := 0; END_IF;
IF Q.Mode <> 1 THEN Q.Motor_RunCmd := FALSE; END_IF;
IF NOT Q.ItemActive OR (Q.Mode = 3) THEN
    Q.D1_ExtendCmd := FALSE;
    Q.D2_ExtendCmd := FALSE;
END_IF;
Q.CompletionPending := Q.CompletionSequence <> CompletionAck;
Q.ReleaseReady := (Q.Mode = 1) AND I.Drive_RunningFB
    AND NOT Q.ItemActive AND NOT Q.CompletionPending AND clearBeams
    AND I.D1_HomeFB AND NOT I.D1_ExtendedFB AND I.D2_HomeFB AND NOT I.D2_ExtendedFB
    AND I.Runout_Ready;
Q.StackLight_Red := Q.Mode = 3;
Q.StackLight_Green := Q.Mode = 1;
CASE Q.Mode OF
    0: Q.ModeText := 'Stopped';
    1: Q.ModeText := 'Auto';
    2: Q.ModeText := 'Stopping';
    3: Q.ModeText := 'Faulted';
END_CASE;
prev := I;

METHOD PRIVATE Finish
VAR_INPUT
    Actual : UINT;
    Result : UINT;
END_VAR
IF Q.ItemActive THEN
    Q.ActualExit := Actual;
    Q.Disposition := Result;
    Q.CompletionSequence := Q.CompletionSequence + 1;
    Q.CompletionItemId := Q.ActiveItemId;
    Q.CompletionRoute := Q.RequestedRoute;
    Q.CompletionExit := Actual;
    Q.CompletionDisposition := Result;
    CASE Actual OF
        1: Q.CountExitA := Q.CountExitA + 1;
        2: Q.CountExitB := Q.CountExitB + 1;
        3: Q.CountRunout := Q.CountRunout + 1;
    END_CASE;
    IF Result = 3 THEN
        Q.CountMisroute := Q.CountMisroute + 1;
        Q.ExceptionCode := 2;
        Q.ExceptionText := 'Misroute: observed exit differs from requested route';
    END_IF;
    IF Result = 4 THEN Q.CountFaulted := Q.CountFaulted + 1; END_IF;
    Q.ItemActive := FALSE;
END_IF;
END_METHOD

METHOD PRIVATE Trip
VAR_INPUT
    Code : UINT;
    Text : STRING(80);
END_VAR
IF Q.Mode <> 3 THEN
    Q.FaultCode := Code;
    Q.FaultText := Text;
    Q.Mode := 3;
    Finish(Actual := 0, Result := 4);
END_IF;
END_METHOD
END_FUNCTION_BLOCK

(* ---- PLC_PRG.st ---- *)
PROGRAM PLC_PRG
VAR
    BenchIntercept : FB_BenchIntercept;
    Conveyor : FB_DemoConveyor;
END_VAR
// First call latches one complete raw image for all downstream application logic.
BenchIntercept(Hardware := GVL_DemoHardware.Inputs);
Conveyor(I := BenchIntercept.Image, NowUs := GVL_BenchRead.PlcTimeUs,
    StartSequence := GVL_DemoWrite.StartSequence,
    StopSequence := GVL_DemoWrite.StopSequence,
    ResetSequence := GVL_DemoWrite.ResetSequence,
    AutoRequest := GVL_DemoWrite.AutoRequest,
    OfferSequence := GVL_DemoWrite.OfferSequence,
    OfferItemId := GVL_DemoWrite.OfferItemId,
    OfferRoute := GVL_DemoWrite.OfferRoute,
    CompletionAck := GVL_DemoWrite.CompletionAck);
GVL_DemoRead.Status := Conveyor.Q;

// Authentic application commands, tapped before the physical sink.
GVL_BenchRead.Motor_RunCmd := Conveyor.Q.Motor_RunCmd;
GVL_BenchRead.D1_ExtendCmd := Conveyor.Q.D1_ExtendCmd;
GVL_BenchRead.D2_ExtendCmd := Conveyor.Q.D2_ExtendCmd;
GVL_BenchRead.StackLight_Red := Conveyor.Q.StackLight_Red;
GVL_BenchRead.StackLight_Green := Conveyor.Q.StackLight_Green;
GVL_DemoHardware.Motor_RunCmd := Conveyor.Q.Motor_RunCmd;
GVL_DemoHardware.D1_ExtendCmd := Conveyor.Q.D1_ExtendCmd;
GVL_DemoHardware.D2_ExtendCmd := Conveyor.Q.D2_ExtendCmd;
GVL_DemoHardware.StackLight_Red := Conveyor.Q.StackLight_Red;
GVL_DemoHardware.StackLight_Green := Conveyor.Q.StackLight_Green;
GVL_BenchRead.OutputSourceEpoch := GVL_BenchRead.AppliedEpoch;
GVL_BenchRead.OutputSourceSequence := GVL_BenchRead.AppliedSequence;
GVL_BenchRead.OutputSourceAppliedCycle := GVL_BenchRead.AppliedCaptureCycle;
GVL_BenchRead.OutputCaptureCycle := GVL_BenchRead.PlcCycle;
GVL_BenchRead.OutputCaptureTimeUs := GVL_BenchRead.PlcTimeUs;
END_PROGRAM
